(* Schneider Machine Expert - Basic project modbus_05_write_single_coil_fc5, file version 3.0.0.0 *)
(* ProjectInformations: Name=New project *)

HARDWARE
  Cpu 0: TM200CE40T
  EthernetConfiguration: NetworkName=M200, IpAllocationMode=FixedAddress, IpAddress=0.0.0.0, SubnetMask=0.0.0.0
  SerialLineConfiguration: Baud=Baud19200, Parity=ParityEven, DataBits=DataBits8, StopBits=StopBits1, PhysicalMedium=PhysicalMediumRs485, TransmissionMode=TransmissionModeModbusRtu, SlaveId=1, Addressing=MasterAddressing
  MastTask: UsePeriodScanMode=false, PeriodScan=100
  FastTask: Period=255
  CpuBehavior: StartingMode=StartAsPreviousState, AutoSaveRamOnEeprom=true, WatchdogPeriod=250

SYMBOLS  (address, symbol, comment, settings)
  %WRITE_VAR0   [Link(Value(FBComLinkParameterEnums=SerialLine1)), RemoteDeviceId(Value(int=1)), Timeout(Value(int=100)), ObjType(Value(FBComObjTypeParameterEnums=SINGLE_COIL)), FirstObj(Value(int=107)), Quantity(Value(int=1)), IndexData(Value(int=260))]

POU Generated C++ - EXPERIMENTAL
  (* SectionNumber=0 *)

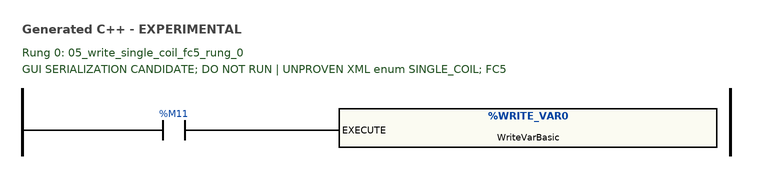

// Rung 0: 05_write_single_coil_fc5_rung_0
// GUI SERIALIZATION CANDIDATE; DO NOT RUN | UNPROVEN XML enum SINGLE_COIL; FC5
  BLK %WRITE_VAR0
  LD %M11
  EXECUTE
  END_BLK
  // as ST:
  //   %WRITE_VAR0(EXECUTE := %M11);
